{region 'Documentation'}
(*!
<summary>Check that the token count is greater than Minimum.</summary>
<description>

StartIndex is an absolute declared IN index, not an offset. Length selects 1..255
elements; the complete selected range must fit IN. Invalid references or ranges report
Error.

Keep supplied arrays stable for the call. Input data is read, not copied or retained as a
snapshot.

Comparison applies Mask to both values; bits outside it are ignored. The default mask
selects all bits.

Counts the currently selected region on evaluation, not occurrences across cycles.
TokenCount exposes the last computed count.

The value token matches under Mask; bits outside Mask are ignored.

</description>
*)
{endregion}
FUNCTION_BLOCK AssertValueTokenCntGreaterThan_Word EXTENDS AssertionBase
VAR_INPUT
    StartIndex : DINT; //! First selected index in IN; uses the array's declared index range, not a zero-based offset.
    Length : USINT; //! Number of selected elements starting at StartIndex; must fit the array range; valid range 1..255.
    Minimum : UINT; //! Exclusive lower bound; the actual value or count must be greater.
    Token : WORD; //! Value searched for in the selected range; Mask selects the compared bits.
    Mask : WORD := WORD#16#FFFF; //! Bits included in the comparison; bits outside the mask are ignored.
END_VAR
VAR_IN_OUT CONSTANT
    IN : ARRAY[*] OF WORD; //! Keep the searched data stable during the call.
END_VAR
VAR
    FTokenCount : UINT;
END_VAR

SUPER^();

{region 'Documentation'}
(*!
<summary>Validate configuration, count tokens and apply the count predicate.</summary>
*)
{endregion}
METHOD PROTECTED Assert
VAR
    InLowerIndex : DINT;
    InUpperIndex : DINT;
    EndIndex : LINT;
    Message : STRING(GVL_Constants.MessageLength);
END_VAR
VAR CONSTANT
    HexDigitCount : USINT := 4;
END_VAR
IF NOT EvaluationActive THEN
    RETURN;
END_IF;

IF Result = E_Result.Error THEN
    RETURN;
END_IF;

// C0371: FB input is checked before any reference access.
{warning disable C0371}
IF NOT __ISVALIDREF(IN) THEN
    FTokenCount := 0;
    Error(Message := 'Assertion error: IN reference is invalid.');
    RETURN;
END_IF;

InLowerIndex := LOWER_BOUND(IN, 1);
InUpperIndex := UPPER_BOUND(IN, 1);
EndIndex := DINT_TO_LINT(StartIndex) + USINT_TO_LINT(Length) - 1;
IF (Length = 0)
    OR (StartIndex < InLowerIndex) OR (StartIndex > InUpperIndex)
    OR (EndIndex > DINT_TO_LINT(InUpperIndex)) THEN
    FTokenCount := 0;
    Message := CONCAT('Assertion error: invalid search range. StartIndex = ',
        DINT_TO_STRING(StartIndex));
    Message := CONCAT(Message, ', Length = ');
    Message := CONCAT(Message, USINT_TO_STRING(Length));
    Error(Message := Message);
    RETURN;
END_IF;

IF Result = E_Result.Failed THEN
    RETURN;
END_IF;

FTokenCount := CountValueTokens_Word(StartIndex := StartIndex,
    Length := Length,
    Token := Token,
    Mask := Mask,
    IN := IN);

IF FTokenCount <= Minimum THEN
    Message := CONCAT('Assertion failed: value token count violates GreaterThan. Actual = ',
        UINT_TO_STRING(FTokenCount));
    Message := CONCAT(Message, ', Minimum = ');
    Message := CONCAT(Message, UINT_TO_STRING(Minimum));
    Message := CONCAT(Message, ', Token = ');
    Message := CONCAT(Message, CreateAssertionTextValue_Hex(Value := WORD_TO_LWORD(Token),
        DigitCount := HexDigitCount));
    Message := CONCAT(Message, ', Mask = ');
    Message := CONCAT(Message, CreateAssertionTextValue_Hex(Value := WORD_TO_LWORD(Mask),
        DigitCount := HexDigitCount));
    Fail(Message := Message);
    RETURN;
END_IF;

Pass();
{warning restore C0371}
END_METHOD

{region 'Documentation'}
(*!
<summary>Clear the retained count on framework reset.</summary>
*)
{endregion}
METHOD PROTECTED ResetAssertion
FTokenCount := 0;
END_METHOD

{region 'Documentation'}
(*!
<summary>Return the most recently evaluated token count.</summary>
<description>

Counts occurrences in one selected array region, not across PLC cycles. Retained while
disabled or after Failed; reset and detected configuration errors clear it. Reading this
property does not search the array.

</description>
*)
{endregion}
{attribute 'monitoring' := 'call'}
PROPERTY PUBLIC TokenCount : UINT //! Return the most recently evaluated token count.
GET // PUBLIC
TokenCount := FTokenCount;
END_GET
END_PROPERTY

END_FUNCTION_BLOCK

(* stored: Version 1.1.0.1
   POU AssertValueTokenCntGreaterThan_Word: Id {7538efae-6f44-47b8-9da1-252e615930e4}, SpecialFunc None
   Folder Internal: Id {e6a206f3-0532-4411-8036-1cbf5bdf7c8d}
   Method Assert: Id {583bcfee-ccd0-4bf2-ad87-489c999ff2fe}
   Method ResetAssertion: Id {86ecdc56-5086-4baa-8ebb-aaf125d7514c}
   Property TokenCount: Id {79552212-2e7f-44b8-8340-db1e011a88e9}
   Get Get: Id {dd234e5d-cd27-4ee0-916b-595145594431} *)
